(* IEC 61131-3 sources: plcassist-cli/packages/volt-lsp-iec/test-corpus/bakon-nano/Device/Plc Logic/Application/Library Manager/L_IPAP_ParameterManagerAccess, 21 files *)

(* ---- GETBOOLEANPROPERTY.fun ---- *)
FUNCTION GETBOOLEANPROPERTY : BOOL
VAR_INPUT
	STKEY : WSTRING;
END_VAR
END_FUNCTION

(* ---- GETCOMPANY.fun ---- *)
FUNCTION GETCOMPANY : WSTRING
END_FUNCTION

(* ---- GETNUMBERPROPERTY.fun ---- *)
FUNCTION GETNUMBERPROPERTY : DINT
VAR_INPUT
	STKEY : WSTRING;
END_VAR
END_FUNCTION

(* ---- GETTEXTPROPERTY.fun ---- *)
FUNCTION GETTEXTPROPERTY : WSTRING
VAR_INPUT
	STKEY : WSTRING;
END_VAR
END_FUNCTION

(* ---- GETTEXTPROPERTY2.fun ---- *)
FUNCTION GETTEXTPROPERTY2 : POINTER TO WSTRING
VAR_INPUT
	STKEY : WSTRING;
END_VAR
END_FUNCTION

(* ---- GETTITLE.fun ---- *)
FUNCTION GETTITLE : WSTRING
END_FUNCTION

(* ---- GETVERSION.fun ---- *)
FUNCTION GETVERSION : VERSION
END_FUNCTION

(* ---- GETVERSIONPROPERTY.fun ---- *)
FUNCTION GETVERSIONPROPERTY : VERSION
VAR_INPUT
	STKEY : WSTRING;
END_VAR
END_FUNCTION

(* ---- L_IPAP_CHECKREADRESULT.fun ---- *)
FUNCTION L_IPAP_CHECKREADRESULT : L_IPAP_REQUEST_STATE
VAR_INPUT
	HREADREQUEST : RTS_IEC_HANDLE;
	PREADBUFFER : POINTER TO BYTE;
	UIBUFFERSIZE : UDINT;
	PREADDATASIZE : POINTER TO UDINT;
	PREADDATATYPE : POINTER TO L_IPAP_DATATYPE;
	PREQUESTRESULT : POINTER TO RTS_IEC_RESULT;
END_VAR
END_FUNCTION

(* ---- L_IPAP_CHECKWRITERESULT.fun ---- *)
FUNCTION L_IPAP_CHECKWRITERESULT : L_IPAP_REQUEST_STATE
VAR_INPUT
	HWRITEREQUEST : RTS_IEC_HANDLE;
	PREQUESTRESULT : POINTER TO RTS_IEC_RESULT;
END_VAR
END_FUNCTION

(* ---- L_IPAP_ERRORHANDLING.fun ---- *)
FUNCTION L_IPAP_ERRORHANDLING : L_IPAP_ERRORID
VAR_INPUT
	EINTERNALERROR : L_IPAP_INTERNALERROR;
END_VAR
END_FUNCTION

(* ---- L_IPAP_SENDREADREQUEST.fun ---- *)
FUNCTION L_IPAP_SENDREADREQUEST : RTS_IEC_HANDLE
VAR_INPUT
	WINDEX : WORD;
	BYSUBINDEX : BYTE;
END_VAR
END_FUNCTION

(* ---- L_IPAP_SENDREADREQUEST_BASEPM.fun ---- *)
FUNCTION L_IPAP_SENDREADREQUEST_BASEPM : RTS_IEC_HANDLE
VAR_INPUT
	WINDEX : WORD;
	BYSUBINDEX : BYTE;
END_VAR
END_FUNCTION

(* ---- L_IPAP_SENDWRITEREQUEST.fun ---- *)
FUNCTION L_IPAP_SENDWRITEREQUEST : RTS_IEC_HANDLE
VAR_INPUT
	WINDEX : WORD;
	BYSUBINDEX : BYTE;
	UIVALUESIZE : UDINT;
	PVALUE : POINTER TO BYTE;
END_VAR
END_FUNCTION

(* ---- L_IPAP_SENDWRITEREQUEST_BASEPM.fun ---- *)
FUNCTION L_IPAP_SENDWRITEREQUEST_BASEPM : RTS_IEC_HANDLE
VAR_INPUT
	WINDEX : WORD;
	BYSUBINDEX : BYTE;
	UIVALUESIZE : UDINT;
	PVALUE : POINTER TO BYTE;
END_VAR
END_FUNCTION

(* ---- L_IPAP_SENDWRITEREQUEST_INTERNAL.fun ---- *)
FUNCTION L_IPAP_SENDWRITEREQUEST_INTERNAL : RTS_IEC_HANDLE
VAR_INPUT
	WINDEX : WORD;
	BYSUBINDEX : BYTE;
	UIVALUESIZE : UDINT;
	PVALUE : POINTER TO BYTE;
END_VAR
END_FUNCTION

(* ---- GLOBALTEXTLIST.fb ---- *)
FUNCTION_BLOCK GLOBALTEXTLIST
VAR
	M_TEXTLISTFILE : STRING(255);
	_STNAMESPACE : STRING;
END_VAR
END_FUNCTION_BLOCK

(* ---- IMAGEPOOL.fb ---- *)
FUNCTION_BLOCK IMAGEPOOL
VAR
	M_STNAMESPACE : STRING(80);
	M_STHELPVARID : STRING;
	M_STHELPVARPATH : STRING(255);
	M_STHELP : STRING;
	M_REGISTERIMAGES : BOOL := TRUE;
END_VAR
END_FUNCTION_BLOCK

METHOD FB_INIT : BOOL
VAR_INPUT
	BINITRETAINS : BOOL;
	BINCOPYCODE : BOOL;
END_VAR
END_METHOD

METHOD FB_REINIT : BOOL
END_METHOD

METHOD FB_EXIT : BOOL
VAR_INPUT
	BINCOPYCODE : BOOL;
END_VAR
END_METHOD

(* ---- L_IPAP_CHANGEHTTPSREDIRECTSETTING4EASYUI.fb ---- *)
FUNCTION_BLOCK L_IPAP_CHANGEHTTPSREDIRECTSETTING4EASYUI
VAR_INPUT
	XEXECUTE : BOOL;
	XABORT : BOOL;
	EHTTPSREDIRECTSETTING : L_IPAP_HTTPSREDIRECT;
	UDITIMEOUT : UDINT := 0;
END_VAR
VAR_OUTPUT
	XDONE : BOOL;
	XBUSY : BOOL;
	XABORTED : BOOL;
	XERROR : BOOL;
	EERRORID : L_IPAP_ERRORID;
END_VAR
VAR
	FB_TIMEOUT : TON;
	XEXECUTELAST : BOOL;
	XABORTLAST : BOOL;
	BRESETOUTPUT : BOOL;
	BFALLINGEXECUTE : BOOL;
	BFALLINGABORT : BOOL;
	FBSTATE : L_IPAP_FBSTATE;
	MINDEX : WORD;
	MSUBINDEX : BYTE;
	MSETTING : L_IPAP_HTTPSREDIRECT;
	MREQUESTHANDLE : RTS_IEC_HANDLE;
	MREQUESTSTATE : L_IPAP_REQUEST_STATE;
	MREQUESTRESULT : L_IPAP_INTERNALERROR;
	CURSETTING : USINT;
	UDIDATAREAD : UDINT;
	EDATATYPE : L_IPAP_DATATYPE;
END_VAR
END_FUNCTION_BLOCK

(* ---- L_IPAP_PARAMETERREAD.fb ---- *)
FUNCTION_BLOCK L_IPAP_PARAMETERREAD
VAR_INPUT
	XEXECUTE : BOOL;
	XABORT : BOOL;
	XBASEPARAMETER : BOOL := FALSE;
	WINDEX : WORD;
	BYSUBINDEX : BYTE;
	UDITIMEOUT : UDINT := 0;
	PDATABUFFER : POINTER TO BYTE := 0;
	UDIBUFFERSIZE : UDINT := 0;
END_VAR
VAR_OUTPUT
	XDONE : BOOL;
	XBUSY : BOOL;
	XABORTED : BOOL;
	XERROR : BOOL;
	EERRORID : L_IPAP_ERRORID;
	UDIDATAREAD : UDINT;
	EDATATYPE : L_IPAP_DATATYPE;
END_VAR
VAR
	FB_TIMEOUT : TON;
	XEXECUTELAST : BOOL;
	XABORTLAST : BOOL;
	BRESETOUTPUT : BOOL;
	BFALLINGEXECUTE : BOOL;
	BFALLINGABORT : BOOL;
	FBSTATE : L_IPAP_FBSTATE;
	MREQUESTHANDLE : RTS_IEC_HANDLE;
	MREQUESTSTATE : L_IPAP_REQUEST_STATE;
	MREQUESTRESULT : L_IPAP_INTERNALERROR;
END_VAR
END_FUNCTION_BLOCK

(* ---- L_IPAP_PARAMETERWRITE.fb ---- *)
FUNCTION_BLOCK L_IPAP_PARAMETERWRITE
VAR_INPUT
	XEXECUTE : BOOL;
	XABORT : BOOL;
	XBASEPARAMETER : BOOL := FALSE;
	WINDEX : WORD;
	BYSUBINDEX : BYTE;
	UDITIMEOUT : UDINT := 0;
	PDATABUFFER : POINTER TO BYTE := 0;
	UDIDATASIZE : UDINT := 0;
END_VAR
VAR_OUTPUT
	XDONE : BOOL;
	XBUSY : BOOL;
	XABORTED : BOOL;
	XERROR : BOOL;
	EERRORID : L_IPAP_ERRORID;
END_VAR
VAR
	FB_TIMEOUT : TON;
	XEXECUTELAST : BOOL;
	XABORTLAST : BOOL;
	BRESETOUTPUT : BOOL;
	BFALLINGEXECUTE : BOOL;
	BFALLINGABORT : BOOL;
	FBSTATE : L_IPAP_FBSTATE;
	MREQUESTHANDLE : RTS_IEC_HANDLE;
	MREQUESTSTATE : L_IPAP_REQUEST_STATE;
	MREQUESTRESULT : L_IPAP_INTERNALERROR;
END_VAR
END_FUNCTION_BLOCK
